Fanuc KAREL source: KO00030.KL

PROGRAM KO00030
%NOLOCKGROUP
VAR
  P1: JOINTPOS
  P2: JOINTPOS
  P3: JOINTPOS
  P4: JOINTPOS
  OUT: XYZWPR
BEGIN
  OUT = FRAME(P1, P2, P3, P4)
END KO00030
